(* IEC 61131-3 sources: JingjiangMoonbox/Application/Application/任务列表/Main_Task/套色调整/套色新算法, 4 files *)

(* ---- KS_ArcAxisReachRange.st ---- *)
(*@CES
Name=KS_ArcAxisReachRange
Type=FunctionBlock
TypeGuid=6f9dac99-8de1-4efc-8465-68ac443b7d08
Guid=66d8455d-5d38-4db4-a051-65983b6f267b
HasDeclaration=True
HasImplementation=True
*)
{DECLARATION}
FUNCTION KS_ArcAxisReachRange : BOOL(*套色单轴误差到达阈值内*)
(*置位后就不再复位除非关闭使能*)
VAR_INPUT
	i_xEn:BOOL;(*处理使能*)
	i_byArcId:BYTE;(*套色的ID*)
	i_byArcErr_Threshold:BYTE:=50;(*套色误差阈值@单位丝*)
	i_byContinuousCycleCnt:BYTE:=10;(*持续的圈数@持续这么多幅误差都在阈值以内就认为可以输出标志*)
	i_xArcErrValid:BOOL;(*误差有效标志@误差有效才能比较 否者等等吧*)
	i_iArcErr:INT;(*套色误差值(在让料头未到达的时候误差值写成最大值)*)
	i_pbyCycleCnt:POINTER TO BYTE;(*满足条件后的圈数计数值*)
	i_pxArcReachRangeFlag:POINTER TO BOOL;(*套色到达阈值标志*)
END_VAR
VAR
	iN: INT;
	byArcErr_Threshold: BYTE;(*丝单位*)
	byContinuousCycleCnt: BYTE;(*持续的幅数计数值*)
	xArcReachRangeFlag:BOOL;(*套色到达阈值标志*)
	byCycleCnt:BYTE;(*每个轴的循环计数*)
	iArcErr:INT;(*套色误差*)
END_VAR
VAR_INPUT
END_VAR
VAR
END_VAR

{IMPLEMENTATION}
IF i_pxArcReachRangeFlag<>0 THEN
	xArcReachRangeFlag:=i_pxArcReachRangeFlag^;
END_IF
IF i_pbyCycleCnt<>0 THEN
	byCycleCnt:=i_pbyCycleCnt^;
END_IF

(*阈值参数*)
byArcErr_Threshold:=i_byArcErr_Threshold;
IF byArcErr_Threshold<=0 THEN
	byArcErr_Threshold:=50;
END_IF

(*持续的幅数参数*)
byContinuousCycleCnt:=i_byContinuousCycleCnt;
IF byContinuousCycleCnt=0 THEN
	byContinuousCycleCnt:=10;
END_IF
iArcErr:=i_iArcErr;

IF i_xEn THEN
	IF i_byArcId>=2 AND i_byArcId<=16 THEN(*从2色开始到最后|检查误差值是否在阈值范围以内*)
		IF NOT xArcReachRangeFlag THEN
			IF i_xArcErrValid THEN
				IF ABS(iArcErr)<=byArcErr_Threshold THEN(*在范围内*)
					byCycleCnt:=byCycleCnt+1;
				ELSE(*有一次跳出，就清零*)
					byCycleCnt:=0;
				END_IF
			ELSE(*等等吧*);
			END_IF

			(*检查是否足够设定的幅数@*)
			IF byCycleCnt>byContinuousCycleCnt THEN
				xArcReachRangeFlag:=TRUE;
			END_IF
		ELSE;
		END_IF
	ELSE
		xArcReachRangeFlag:=FALSE;
		byCycleCnt:=0;
	END_IF
ELSE
	(*复位参数*)
	xArcReachRangeFlag:=FALSE;
	byCycleCnt:=0;
END_IF

IF i_pxArcReachRangeFlag<>0 THEN
	i_pxArcReachRangeFlag^:=xArcReachRangeFlag;
END_IF
IF i_pbyCycleCnt<>0 THEN
	i_pbyCycleCnt^:=byCycleCnt;
END_IF

(* ---- KS_ArcCompensate_Hor.st ---- *)
(*@CES
Name=KS_ArcCompensate_Hor
Type=FunctionBlock
TypeGuid=6f9dac99-8de1-4efc-8465-68ac443b7d08
Guid=22f1b56e-db40-40dc-a19f-6fb25d07bc3f
HasDeclaration=True
HasImplementation=True
*)
{DECLARATION}
FUNCTION KS_ArcCompensate_Hor : BOOL
(*套色的横向补偿@针对裁切后横向跑出波门位置丢失*)
VAR_INPUT
	i_xEn					:BOOL;(*补偿使能*)
	i_xDirRev				:BOOL;(*方向取反@默认是误差和调整量同向*)
	i_xCut_Uw				:BOOL;(*裁切标志@放料*)
	i_xCut_Rw				:BOOL;(*裁切标志@收料*)
	i_xLost					:BOOL;(*丢失标志*)
	i_byOutEnLostNum		:BYTE;(*丢失次数@超过该值认为需要补偿输出*)
	i_byAddValue			:BYTE;(*叠加的调整量@丝*)
	i_byMaxAddValue_Total	:BYTE;(*叠加的最大调整量@mm*)
	i_iAdjValue				:INT;(*横向调整量*)
	i_iArcErr				:INT;(*横向误差*)
	i_iMaxAdjustVal			:INT;(*横向最大调整量@um*)
	i_iMinArcErr_Compensate	:INT;(*横向补偿启用的最小误差@丝*)
	i_paiAdjValueList		:POINTER TO ARRAY [1..10] OF INT;(*10幅调整量列表@[10]最新*)
	i_paiArcErrList			:POINTER TO ARRAY [1..10] OF INT;(*10幅套色误差列表@[10]最新*)
	i_pxWatching			:POINTER TO BOOL;(*监控中标志*)
	i_pxOuting				:POINTER TO BOOL;(*输出中标志*)
	i_pxOutDne				:POINTER TO BOOL;(*输出完成*)
	i_pbyLostCnt			:POINTER TO BYTE;(*丢失次数*)
	i_prResult_Total		:POINTER TO REAL;(*总的补偿值@mm*)
	i_prResult				:POINTER TO REAL;(*输出补偿结果值@um*)
END_VAR
VAR
	aiAdjValueList		:ARRAY [1..10] OF INT;(*10幅调整量列表@[10]最新*)
	aiArcErrList		:ARRAY [1..10] OF INT;(*10幅套色误差列表@[10]最新*)
	xWatching			:BOOL;(*监控中标志*)
	xOuting				:BOOL;(*输出中标志*)
	xOutDne				:BOOL;(*输出完成*)
	byLostCnt			:BYTE;(*丢失次数*)
	rResult_Total		:REAL;(*总的补偿值@mm*)
	rResult				:REAL;(*输出补偿结果值@um*)
	iN					:INT;
	iDelta				:INT;
	iNum0				:INT;
	iNum1				:INT;
	rSum				:REAL;
	iCoeff				:INT;(*方向系数*)
	xGTMinArcErr		:BOOL;(*大于最小误差标志@有效了可以输出补偿*)
END_VAR
{IMPLEMENTATION}
IF i_prResult_Total<>0 THEN
	rResult_Total:=i_prResult_Total^;(*重新统计的时候再清除*)
END_IF
IF i_xEn THEN
	(*放到en的好处就是else会直接清除这些变量*)
	IF i_paiAdjValueList<>0 THEN
		aiAdjValueList:=i_paiAdjValueList^;
	END_IF
	IF i_paiArcErrList<>0 THEN
		aiArcErrList:=i_paiArcErrList^;
	END_IF
	IF i_pxWatching<>0 THEN
		xWatching:=i_pxWatching^;
	END_IF
	IF i_pxOuting<>0 THEN
		xOuting:=i_pxOuting^;
	END_IF
	IF i_pxOutDne<>0 THEN
		xOutDne:=i_pxOutDne^;
	END_IF
	IF i_pbyLostCnt<>0 THEN
		byLostCnt:=i_pbyLostCnt^;
	END_IF

	IF i_xCut_Uw AND NOT xWatching THEN(*裁切标志有效@c初始化参数*)
		xWatching:=TRUE;
		xOuting:=FALSE;
		xOutDne:=FALSE;
		byLostCnt:=0;
		rResult_Total:=0;(*清零统计值*)
		FOR iN:=1 TO 10 BY 1 DO
			aiAdjValueList[iN]:=0;
			aiArcErrList[iN]:=0;
		END_FOR
	END_IF

	IF xWatching THEN
		IF i_xLost THEN
			IF byLostCnt<i_byOutEnLostNum THEN
				byLostCnt:=byLostCnt+1;
			ELSE
				xOuting:=TRUE;
			END_IF
		ELSE(*未丢失*)
			byLostCnt:=0;(*重新统计@只要有正常的就重新统计*)
			(*更新误差和调整量列表*)
			KS_PushValueToList(i_iAdjValue, 10, TYPE_INT, ADR(aiAdjValueList));
			KS_PushValueToList(i_iArcErr, 10, TYPE_INT, ADR(aiArcErrList));
		END_IF

		IF xOuting THEN(*计算一次*)
(*
			(*计算调整量方向*)
			(*看前6个点|5个变化量*)
			iNum:=0;
			FOR iN:=10 TO 6 BY -1 DO
				iDelta:=aiArcErrList[iN]-aiArcErrList[iN-1];
				IF iDelta>=0 THEN(*=0 也算有效*)
					iNum:=iNum+1;
				ELSIF iDelta<0 THEN
					iNum:=iNum-1;
				END_IF
			END_FOR

			IF ABS(iNum)>=3 THEN(*50%的数据都是朝一个方向的|我们触发输出*);
			ELSE
				xOuting:=FALSE;
				xOutDne:=TRUE;(*就直接结束吧*)
			END_IF
*)
			xWatching:=FALSE;(*不再监控了*)
			byLostCnt:=0;
		END_IF
	END_IF

	(*输出中*)
	IF xOuting THEN
		(*计算调整量方向*)
		(*看前6个点|5个变化量*)
		iNum0:=0;
		iNum1:=0;
		xGTMinArcErr:=FALSE;
		FOR iN:=10 TO 6 BY -1 DO
			iDelta:=aiArcErrList[iN]-aiArcErrList[iN-1];
			IF iDelta>0 THEN
				iNum0:=iNum0+1;
			ELSIF iDelta<0 THEN
				iNum1:=iNum1+1;
			ELSE;
			END_IF

			(*2024.8.6.172305+误差队列中的误差存在比最小值大的就可以输出补偿*)
			(*用于弥补误差不大的时候由于色标信号消失引起的误动作*)
			IF ABS(aiArcErrList[iN])>i_iMinArcErr_Compensate THEN
				xGTMinArcErr:=TRUE;
			END_IF
		END_FOR

		IF xGTMinArcErr THEN(*有大于最小误差值的*)
			IF iNum0 > iNum1 THEN(*正的多*)
				iCoeff:=1;
			ELSIF iNum0 < iNum1 THEN(*负的多*)
				iCoeff:=-1;
			ELSE(*这次退出*)
				iCoeff:=0;
				xOuting:=FALSE;
				xOutDne:=TRUE;(*就直接结束吧*)
			END_IF
		ELSE(*没有则退出不补偿@省的误动作*)
			iCoeff:=0;
			xOuting:=FALSE;
			xOutDne:=TRUE;(*就直接结束吧*)
		END_IF

		(*计算补偿量*)
		IF FALSE THEN
			(*计算累计调整量的方向作为我补偿的方向*)
			rSum:=0;
			FOR iN:=1 TO 10 BY 1 DO
				rSum:=rSum+aiAdjValueList[iN];
			END_FOR
			IF rSum>0 THEN
				rResult:=BYTE_TO_REAL(i_byAddValue)*10;(*um值*)
			ELSIF rSum<0 THEN
				rResult:=-BYTE_TO_REAL(i_byAddValue)*10;(*um值*)
			ELSE
				rResult:=0;(*um值*)
			END_IF
		ELSE
			rResult:=BYTE_TO_REAL(i_byAddValue)*10;(*um值*)
			rResult:=iCoeff*rResult;
			IF i_xDirRev THEN
				rResult:=-rResult;
			END_IF
		END_IF

		(*做单圈最大输出限制@2024.8.4.195257*)
		IF rResult<>0 THEN
			IF ABS(rResult)>ABS(i_iMaxAdjustVal) THEN
				rResult:=i_iMaxAdjustVal*rResult/ABS(rResult);
			END_IF
		END_IF

		(*检查丢失状态*)
		IF NOT i_xLost THEN(*连续2幅未丢失则交给自动*)
			byLostCnt:=byLostCnt+1;
		END_IF

		rResult_Total:=rResult_Total+rResult;(*累加*)
		IF ABS(rResult_Total)/1000>=i_byMaxAddValue_Total OR
			byLostCnt>=2 THEN(*连续2幅未丢失就结束,则交给自动@byLostCnt 这里做未丢失统计数目使用*)
			xOuting:=FALSE;
			xOutDne:=TRUE;
		END_IF
	END_IF

	(*收料裁切就强制结束*)
	IF i_xCut_Rw THEN
		xOuting:=FALSE;
		xOutDne:=TRUE;
		xWatching:=FALSE;(*不再监控了*)
	END_IF
ELSE;
END_IF

IF i_paiAdjValueList<>0 THEN
	i_paiAdjValueList^:=aiAdjValueList;
END_IF
IF i_paiArcErrList<>0 THEN
	i_paiArcErrList^:=aiArcErrList;
END_IF
IF i_pxWatching<>0 THEN
	i_pxWatching^:=xWatching;
END_IF
IF i_pxOuting<>0 THEN
	i_pxOuting^:=xOuting;
END_IF
IF i_pxOutDne<>0 THEN
	i_pxOutDne^:=xOutDne;
END_IF
IF i_pbyLostCnt<>0 THEN
	i_pbyLostCnt^:=byLostCnt;
END_IF
IF i_prResult_Total<>0 THEN
	i_prResult_Total^:=rResult_Total;
END_IF
IF i_prResult<>0 THEN
	i_prResult^:=rResult;
END_IF

(* ---- KS_GetArcKAdjBySts.st ---- *)
(*@CES
Name=KS_GetArcKAdjBySts
Type=FunctionBlock
TypeGuid=6f9dac99-8de1-4efc-8465-68ac443b7d08
Guid=ab0b9e35-35e9-482c-8b4f-391e87029d49
HasDeclaration=True
HasImplementation=True
*)
{DECLARATION}
FUNCTION KS_GetArcKAdjBySts : BYTE
(*2024.9.2.104007*)
(*根据套色调整状态输出增益,@=0 初始状态(增益略大) |=1 稳态状态(增益略小)*)
(*匀速,速度高于一定值才判断,反之使用初始误差,
连续一定幅最多20幅误差小于一定值,变化量也小于一定值认为稳态*)
(*2024.9.6.124942 增加计算*)
VAR_INPUT
	i_xEn						: BOOL;(*使能标志@未使能则使用初始增益*)
	i_byKadj_SetType			: BYTE;(*套色K值设置方式
								@ =0 使用初始增益|计算Ki的速度=当前速度@实际积分的系数是定值
								@ =1 使用初始增益的同时,计算Ki的速度也是定值-按照30m/min输出@实际积分的系数是随速度减小的
								@ =2 根据状态设置|计算Ki的速度根据当前速度变化@实际积分的系数是定值
								@ =3 根据状态设置的同时,计算Ki的速度也是定值-按照30m/min输出@实际积分的系数是随速度减小的*)
	i_rKadj_PID_Mol_Init 		: REAL;(*模型的pid增益_初始增益@开机和接料使用*)
	i_rKadj_I_Mol_Init			: REAL;(*模型的I值增益_初始增益@开机和接料使用*)
	i_rKadj_PID_Mol_SteadySts	: REAL;(*模型的pid增益_稳态增益*)
	i_rKadj_I_Mol_SteadySts		: REAL;(*模型的I值增益_稳态增益*)
	i_xCut						: BOOL;(*裁切了@沿标志|判定状态使用*)
	i_xFilmArrived_Cut			: BOOL;(*裁切后料膜到达@让料头标志*)
	i_xEvenning					: BOOL;(*匀速状态@此时才能判定状态*)
	i_iVel_Cur					: INT;(*当前速度@m/min*)
	i_iErrValue					: INT;(*误差值@丝*)
	i_byErrThreshold			: BYTE:=30;(*套色误差阈值@单位丝|判定状态使用*)
	i_byDeltaErrThreshold		: BYTE:=10;(*套色误差变化量阈值@单位丝|判定状态使用*)
	i_iVelThreshold				: INT:=100;(*速度阀值@超过该速度才判断状态@允许=0*)

	i_pxCutting					: POINTER TO BOOL;(*裁切中标志*)
	i_paiErrValueList			: POINTER TO ARRAY [0..20] OF INT;(*20个缓存[20]=最新值@[0]=统计缓存个数*)
	i_pbyArcAdjSts				: POINTER TO BYTE;(*套色调整状态@=0 初始状态(增益略大) |=1 稳态状态(增益略小)*)
	i_prKadj_Pid				: POINTER TO REAL;(*输出的增益值*)
	i_prKadj_I					: POINTER TO REAL;(*输出的增益值*)
	i_prVel_Ki					: POINTER TO REAL;(*计算的ki的速度@2024.9.6.123736根据状态会变化*)
END_VAR
VAR
	rKadj_Pid				: REAL;(*输出的增益值*)
	rKadj_I					: REAL;(*输出的增益值*)
	xUseInitKAdj			: BOOL:=TRUE;(*默认使用初始k|反之则使用状态k*)
	byArcAdjSts				: BYTE;(*套色调整状态*)
	aiErrValueList			: ARRAY [1..20] OF INT;(*20个缓存[20]=最新值*)
	iErrValueListNum		: INT;(*缓存个数*)
	iErrValue				: INT;(*误差值*)
	iDeltaValue				: INT;(*变化量*)
	iErrNum					: INT;(*误差个数*)
	iN						: INT;(*循环*)
	iErrValue1				: INT;(*前一个误差*)
	iErrValue2				: INT;(*较新的误差*)
	xUpdatErrList			: BOOL;(*更新误差列表*)
	iVelThreshold			: INT;(*速度阈值临时*)
	xJudgeAdjSts			: BOOL;(*判断状态标志*)
	xIsSteadySts			: BOOL;(*已经是稳态了*)
	xNotSteadySts			: BOOL;(*s是非稳态@不再判断了*)
	xCutting				: BOOL;(*裁切中*)
	rVel_Ki					: REAL;(*计算Ki的速度*)
END_VAR
{IMPLEMENTATION}
IF i_pxCutting<>0 THEN
	xCutting:=i_pxCutting^;
END_IF

IF i_paiErrValueList<>0 THEN
	iErrValueListNum:=i_paiErrValueList^[0];
	SysMemCpy(ADR(aiErrValueList),ADR(i_paiErrValueList^[1]),SIZEOF(aiErrValueList));
END_IF
IF i_pbyArcAdjSts<>0 THEN
	byArcAdjSts:=i_pbyArcAdjSts^;
END_IF

iErrValue:=i_iErrValue;
iVelThreshold:=i_iVelThreshold;
iErrNum:=SIZEOF(aiErrValueList)/SIZEOF(aiErrValueList[1]);

IF i_xEn THEN
	IF i_byKadj_SetType = 2 OR i_byKadj_SetType=3 THEN(*根据状态切换增益*)
		xUseInitKAdj:=FALSE;
		(*裁切状态切换*)
		IF i_xCut THEN
			xCutting:=TRUE;
		ELSIF xCutting THEN
			IF i_xFilmArrived_Cut THEN
				xCutting:=FALSE;
			END_IF
		END_IF

		(*套色误差判断状态*)
		IF iErrValueListNum	< iErrNum THEN
			byArcAdjSts:=0;
			iErrValueListNum:=iErrValueListNum+1;(*开始累*)
			aiErrValueList[iErrValueListNum] := i_iErrValue;
		ELSE
			xUpdatErrList:=TRUE;
		END_IF

		(*判断是否已经进入了稳态*)
		IF byArcAdjSts=1 THEN
			xIsSteadySts:=TRUE;
		END_IF

		IF iErrValueListNum>= iErrNum THEN(*累计足够了*)
			FOR iN:=1 TO iErrNum-1 BY 1 DO
				(*更新列表*)
				IF xUpdatErrList THEN
					IF iN=1 THEN(*直接更新[1] [2],这样下面的计算才正确*)
						aiErrValueList[iN] := aiErrValueList[iN+1];
						aiErrValueList[iN+1] := aiErrValueList[iN+2];
					ELSIF iN<iErrNum-1 THEN(*=2 更新第3个|以此类推*)
						aiErrValueList[iN+1] := aiErrValueList[iN+2];
					ELSE(*更新最后一个*)
						aiErrValueList[iN+1] := i_iErrValue;
					END_IF
				END_IF

				(*获取误差*)
				iErrValue1:=aiErrValueList[iN];
				iErrValue2:=aiErrValueList[iN+1];
				iDeltaValue:=iErrValue2-iErrValue1;

				xJudgeAdjSts:=i_iVel_Cur>=iVelThreshold AND i_xEvenning;(*高速,匀速,才判断套色状态*)
				xJudgeAdjSts:=xJudgeAdjSts AND NOT xCutting;(*处于非裁切中才进行状态判定*)
				IF xJudgeAdjSts THEN
					IF NOT xIsSteadySts AND NOT xNotSteadySts THEN(*未进入稳态|没有判断出是非稳态*)
						IF iN=1 THEN(*判断2个误差的阈值*)
							IF ABS(iErrValue1)<=i_byErrThreshold AND
								ABS(iErrValue2)<=i_byErrThreshold AND
								ABS(iDeltaValue)<=i_byDeltaErrThreshold THEN
								byArcAdjSts:=1;(*稳态了*)
							ELSE
								byArcAdjSts:=0;(*非稳态了*)
								xNotSteadySts:=TRUE;
							END_IF
						ELSE(*判断较新误差的判断*)
							IF ABS(iErrValue2)<=i_byErrThreshold AND
								ABS(iDeltaValue)<=i_byDeltaErrThreshold THEN
								byArcAdjSts:=1;(*稳态了*)
							ELSE
								byArcAdjSts:=0;(*非稳态了*)
								xNotSteadySts:=TRUE;
							END_IF
						END_IF
					ELSE(*已经进入稳态了*);
					END_IF
				ELSE(*低速都按照初始误差了*)
					byArcAdjSts:=0;(*强制使用初始误差*)
				END_IF
			END_FOR
		END_IF

		IF i_byKadj_SetType=3 THEN(*输出速度为定值*)
			rVel_Ki:=30;
		ELSE(*输出速度根据当前速度变化*)
			rVel_Ki:=i_iVel_Cur;
		END_IF
	ELSE(*使用初始增益*)
		byArcAdjSts:=0;
		xCutting:=FALSE;
		IF iErrValueListNum<>0 THEN
			iErrValueListNum:=0;
			SysMemSet(ADR(aiErrValueList),0,SIZEOF(aiErrValueList));
		END_IF

		IF i_byKadj_SetType=1 THEN(*输出速度为定值*)
			rVel_Ki:=30;
		ELSE(*输出速度根据当前速度变化*)
			rVel_Ki:=i_iVel_Cur;
		END_IF
	END_IF
ELSE
	byArcAdjSts:=0;
	xCutting:=FALSE;
	(*缓存清除*)
	IF iErrValueListNum<>0 THEN
		iErrValueListNum:=0;
		SysMemSet(ADR(aiErrValueList),0,SIZEOF(aiErrValueList));
	END_IF
	rVel_Ki:=i_iVel_Cur;(*按照当前速度输出@2024.9.6.124559*)
END_IF

(*未处理逐步切换*)
IF xUseInitKAdj THEN(*使用初始k*)
	rKadj_Pid:=i_rKadj_PID_Mol_Init;
	rKadj_I:=i_rKadj_I_Mol_Init;
ELSE(*使用状态k*)
	IF byArcAdjSts =1 THEN
		rKadj_Pid:=i_rKadj_PID_Mol_SteadySts;
		rKadj_I:=i_rKadj_I_Mol_SteadySts;
	ELSE
		rKadj_Pid:=i_rKadj_PID_Mol_Init;
		rKadj_I:=i_rKadj_I_Mol_Init;
	END_IF
END_IF

IF i_pbyArcAdjSts<>0 THEN
	i_pbyArcAdjSts^:=byArcAdjSts;
END_IF
IF i_prKadj_Pid<>0 THEN
	i_prKadj_Pid^:=rKadj_Pid;
END_IF
IF i_prKadj_I<>0 THEN
	i_prKadj_I^:=rKadj_I;
END_IF
IF i_pxCutting<>0 THEN
	i_pxCutting^:=xCutting;
END_IF
IF i_paiErrValueList<>0 THEN
	i_paiErrValueList^[0]:=iErrValueListNum;
	SysMemCpy(ADR(i_paiErrValueList^[1]),ADR(aiErrValueList),SIZEOF(aiErrValueList));
END_IF
IF i_prVel_Ki<>0 THEN
	i_prVel_Ki^:=rVel_Ki;
END_IF

(* ---- KS_PushValueToList.st ---- *)
(*@CES
Name=KS_PushValueToList
Type=FunctionBlock
TypeGuid=6f9dac99-8de1-4efc-8465-68ac443b7d08
Guid=e04ac46d-5d6b-4101-9912-eb5ef8957014
HasDeclaration=True
HasImplementation=True
*)
{DECLARATION}
FUNCTION KS_PushValueToList : BOOL
(*将输入值写入到列表|最后一个数据为最新数据|只处理了int类型数据*)
VAR_INPUT
	i_rValue:REAL;(**)
	i_uiDataNum:UINT;(*数据个数*)
	i_iDataType:TypEnumDataType;(*数据类型*)
	i_dwListAdr:DWORD;(*数据的起始地址*)
END_VAR
VAR
	iN: INT;
	piTmp:POINTER TO INT;
	piTmp_Next:POINTER TO INT;
	iDeltaLenth: INT;
END_VAR
{IMPLEMENTATION}
IF i_uiDataNum>0 AND i_dwListAdr<>0 THEN
	CASE i_iDataType OF
		TYPE_INT:
			iDeltaLenth:=2;(*偏移2个字节*)

			piTmp:=i_dwListAdr;
			IF i_uiDataNum<>1 THEN
				FOR iN:=1 TO UINT_TO_INT(i_uiDataNum)-1 BY 1 DO
					piTmp_Next:=piTmp+INT_TO_DWORD(iDeltaLenth);
					piTmp^:=piTmp_Next^;(*将下一个数据写入到当前位置*)
					piTmp:=piTmp+INT_TO_DWORD(iDeltaLenth);
				END_FOR
				piTmp^:=REAL_TO_INT(i_rValue);
			ELSE(*只有一个数据*)
				piTmp^:=REAL_TO_INT(i_rValue);
			END_IF
	ELSE;
	END_CASE

ELSE;
END_IF
